(* IEC 61131-3 sources: plcassist-cli/packages/volt-lsp-iec/test-corpus/bakon-nano/Device/Plc Logic/Application/Library Manager/TextListUtils, 11 files *)

(* ---- GVL_TEXTLISTINFO.gvl ---- *)
VAR_GLOBAL
	FACTORY : TextListInfoFactory;
END_VAR

(* ---- ITEXTLISTINFO.itf ---- *)
INTERFACE ITEXTLISTINFO
END_INTERFACE

METHOD GETIDITERATOR : COL.IIterator
END_METHOD

METHOD RELEASE : BOOL
END_METHOD

(* ---- CREATEADDITIONALELEMENT_CB.fun ---- *)
FUNCTION CREATEADDITIONALELEMENT_CB : BOOL
VAR_INPUT
	PSTID : POINTER TO BYTE;
	PFBTEXTLISTINFO : POINTER TO TextListInfo;
END_VAR
END_FUNCTION

(* ---- GETLANGUAGETEXT.fun ---- *)
FUNCTION GETLANGUAGETEXT : ReturnValues
VAR_INPUT
	PSTEXT : POINTER TO STRING;
	DISIZE : DINT;
END_VAR
VAR_OUTPUT
	BDEFAULTTEXT : BOOL;
END_VAR
VAR_IN_OUT
	STEXTLIST : STRING;
	STEXTINDEX : STRING;
	SLANGUAGE : STRING;
END_VAR
END_FUNCTION

(* ---- GETLANGUAGETEXTW.fun ---- *)
FUNCTION GETLANGUAGETEXTW : ReturnValues
VAR_INPUT
	PWSTEXT : POINTER TO WSTRING;
	DISIZE : DINT;
END_VAR
VAR_OUTPUT
	BDEFAULTTEXT : BOOL;
END_VAR
VAR_IN_OUT
	STEXTLIST : STRING;
	STEXTINDEX : STRING;
	SLANGUAGE : STRING;
END_VAR
END_FUNCTION

(* ---- GETTEXT.fun ---- *)
FUNCTION GETTEXT : ReturnValues
VAR_INPUT
	PSTEXT : POINTER TO STRING;
	DISIZE : DINT;
END_VAR
VAR_OUTPUT
	BDEFAULTTEXT : BOOL;
END_VAR
VAR_IN_OUT
	STEXTLIST : STRING;
	STEXTINDEX : STRING;
END_VAR
END_FUNCTION

(* ---- GETTEXTLISTINFO.fun ---- *)
FUNCTION GETTEXTLISTINFO : ITextListInfo
VAR_IN_OUT
	STTEXTLISTNAME : STRING(255);
END_VAR
END_FUNCTION

(* ---- GETTEXTW.fun ---- *)
FUNCTION GETTEXTW : ReturnValues
VAR_INPUT
	PWSTEXT : POINTER TO WSTRING;
	DISIZE : DINT;
END_VAR
VAR_OUTPUT
	BDEFAULTTEXT : BOOL;
END_VAR
VAR_IN_OUT
	STEXTLIST : STRING;
	STEXTINDEX : STRING;
END_VAR
END_FUNCTION

(* ---- TEXTLISTINFO.fb ---- *)
FUNCTION_BLOCK TEXTLISTINFO EXTENDS InstanceBase
VAR
	M_STEXTLISTNAME : STRING(255);
	M_LISTOFENTRIES : COL.IList;
	M_ITFLISTFACTORY : COL.ListFactory;
	M_STRINGFACTORY : COL.StringElementFactory;
	M_ITERATORFB : COL.ListIterator;
	M_XTEXTLISTREAD : BOOL;
	NAME : STRING(255);
	NUMBEROFENTRIES : UDINT;
END_VAR
END_FUNCTION_BLOCK

METHOD ADDELEMENT : BOOL
VAR_INPUT
	PSTID : POINTER TO STRING(80);
END_VAR
END_METHOD

METHOD PRVINSTINIT : FBF.ERROR
VAR_INPUT
	ITFDATA : FBF.IData;
END_VAR
END_METHOD

METHOD GETIDITERATOR : COL.IIterator
END_METHOD

METHOD RELEASE : BOOL
END_METHOD

(* ---- TEXTLISTINFODATA.fb ---- *)
FUNCTION_BLOCK TEXTLISTINFODATA EXTENDS InstanceData
VAR_INPUT
	STTEXTLISTNAME : STRING(255);
END_VAR
END_FUNCTION_BLOCK

(* ---- TEXTLISTINFOFACTORY.fb ---- *)
FUNCTION_BLOCK TEXTLISTINFOFACTORY EXTENDS FactoryBase
VAR
	PRVINSTCOUNT : CAA.COUNT;
	PRVINSTPOOLEXTENDSFACTOR : USINT;
	PRVINSTSIZE : CAA.SIZE;
END_VAR
END_FUNCTION_BLOCK

METHOD CREATE : ITextListInfo
VAR_INPUT
	STTEXTLISTNAME : STRING(255);
END_VAR
VAR_OUTPUT
	EERROR : FBF.ERROR;
END_VAR
END_METHOD
